(* IEC 61131-3 sources: SRCI_CLIENT_PLC/RobotLibrary/Library/POUs/General/MC_RobotTask/Structures/ParCfg, 1 file *)

(* ---- RobotTaskParCfg.st ---- *)
{attribute 'pack_mode' := '1'}
// -------------------------------------------------------------------------
//  SRCI Robot Library
// -------------------------------------------------------------------------
//
//  Object:      RobotTaskParCfg
//  Author:      Thorsten Brach
//  Date:        2024-11-30
//
//  Description:
//
//
//  Copyright:
//    (C) 2024 Thorsten Brach. All rights reserved
//             Licensed under the MIT License.
//
//  Disclaimer:
//    This project is provided without any guarantee and can be used for
//    private and commercial purposes. Any use is at the user’s
//    own risk and responsibility.
//
// -------------------------------------------------------------------------
TYPE RobotTaskParCfg :
STRUCT
  /// Common parameter
  Com    : RobotTaskParCfgCom;
  /// PLC parameter
  Plc    : RobotTaskParCfgPlc;
  /// Robot parameter
  Rob    : RobotTaskParCfgRob;
END_STRUCT
END_TYPE
